Staubli VAL3: exercice3.pgx

program exercice3()
  local num l_n1
begin
  movej(jDepart,tPince,mRapide)
  call ouvrirPince()

  for l_n1 = 0 to 4
    movej(appro(Prise5[l_n1],{0,0,-50,0,0,0}),tPince,mRapide)
    movel(Prise5[l_n1],tPince,mLent)
    call fermerPince()
    movel(appro(Prise5[l_n1],{0,0,-50,0,0,0}),tPince,mRapide)

    movej(jDepart,tPince,mRapide)
    movej(appro(pDepose[0],{0,0,-50,0,0,0}),tPince,mRapide)
    movel(pDepose[0],tPince,mLent)
    call ouvrirPince()
    movel(appro(pDepose,{0,0,-50,0,0,0}),tPince,mRapide)


    movej(jDepart,tPince,mLent)
    waitEndMove()
    delay(3)
  endFor

end
